(* PLC project Vn_networks_mixed4, Beckhoff Automation GmbH TwinCAT PLC Control 3.5.13.21 *)
(* stored: creationDateTime 1970-01-01T00:00:00 *)

PROGRAM Vn_networks_mixed4

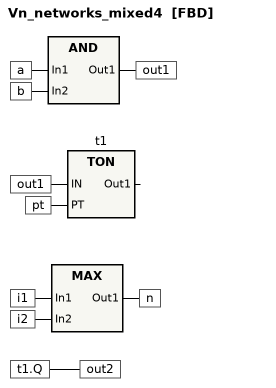
(* FBD diagram, written out as Structured Text *)
out1 := a AND b;
t1(IN := out1, PT := pt);
n := MAX(i1, i2);
out2 := t1.Q;
END_PROGRAM
